(* IEC 61131-3 sources: kns-port-domestic/tools/plcopen/tests/fixtures/constructs/src/POUs/PRG_Aux, 3 files *)

(* ---- PRG_Aux.decl.st ---- *)
// Назначение: программа с методом; комментарии всех видов
// Автор:      <ИМЯ ФАМИЛИЯ>
// Версия:     0.1.0
// Документ:   docs/plcopen.md
PROGRAM PRG_Aux
VAR
    fbValve : FB_Valve;
    itfPos : I_Positioner;
    itfLock : I_Lockable;
    iCalls : INT;
    wsMsg : WSTRING(32) := "Задвижка <закрыта> & 'ok'";
    sMsg : STRING(32) := 'a$'b"c <&>';
END_VAR
VAR_EXTERNAL
    xDoRun : BOOL;              // выход из GVL_Io (необязательное объявление CODESYS)
END_VAR

(* ---- PRG_Aux.impl.st ---- *)
(* внешний (* вложенный *) комментарий *)
itfPos := fbValve;
itfLock := fbValve;
itfPos.Setpoint := 50.0;
itfPos.MoveTo(rPos_pct := 40.0);
itfLock.Lock(xLock := NOT xDoRun);
fbValve();
Step(iInc := 1);
F_Noop(xIn := TRUE);
IF iCalls > 5 AND_THEN fbValve.rPos_pct < 1.0E3 THEN
    iCalls := 0;
END_IF

(* ---- Step.method.decl.st ---- *)
// Шаг программы
METHOD Step : INT
VAR_INPUT
    iInc : INT := 1;
END_VAR
